FUNCTION_BLOCK FB_ReadPressure
VAR_INPUT
	bExecute	:	BOOL	:=	FALSE;
END_VAR
VAR_OUTPUT
	bBusy		:	BOOL	:=	FALSE;
	bErr		:	BOOL	:=	FALSE;
	Pressure	:	REAL	:=	0.0;
END_VAR
VAR
	nState		:	UDINT	:=	0;
END_VAR

// bNordReadAcc 키면서
// busy state로 올림

// press 읽어서 PYADS에 입력하고
// 다 입력되면 NordPress에 쓰고 bNordReadAcc 끄기
// 만약 실패시 busy 끄면서 fail 올리기



CASE nState OF

0:
	IF bExecute	THEN
		PYADSPort.bNordReadReq	:=	TRUE;
		bBusy	:=	TRUE;
		nState	:=	1;
	END_IF

1:
	IF NOT PYADSPort.bNordReadReq THEN
		IF PYADSPort.bNordReadErr THEN
			PYADSPort.bNordReadErr	:=	FALSE;
			bErr	:=	TRUE;
		ELSE
			bErr	:=	FALSE;
		END_IF
			Pressure:=	PYADSPort.nNordPress;
			bBusy	:=	FALSE;
			nState	:=	0;
	END_IF
END_CASE

END_FUNCTION_BLOCK

(* stored: Version 1.1.0.1, ProductVersion 3.1.4024.15
   POU FB_ReadPressure: Id {3eedfdbd-e9c2-4df2-be20-e62e60da9873}, SpecialFunc None *)
